// TIA Portal V18 export
// export: Created 2026-11-18T07:26:10.6281665Z, ExportSetting WithDefaults, DisplayName Totally Integrated Automation Portal, DisplayVersion V18 Update 6, DisplayName TIA Portal Openness, DisplayVersion V18 Update 6, DisplayName TIA Portal Version Control Interface, DisplayVersion V18, DisplayName SINAMICS Startdrive Advanced, DisplayVersion V18 SP2 Update 1, DisplayName SINAMICS DCC, DisplayVersion V18 Update 1, DisplayName SINAMICS Startdrive G110M, G120, G120C, G120D, G120P, G115D, DisplayVersion V18 SP2 Update 1, DisplayName SINAMICS Startdrive G130, G150, S120, S150, SINAMICS MV, S210, G220, S200, DisplayVersion V18 SP2 Update 1, DisplayName STEP 7 Professional, DisplayVersion V18 Update 6, DisplayName STEP 7 CFC, DisplayVersion V18 Update 2, DisplayName STEP 7 Safety, DisplayVersion V18, DisplayName WinCC Professional, DisplayVersion V18 Update 6
PlcWatchTable "Drive_1_Izleme"
  PlcWatchTableEntry ""Motor1_Start""  DisplayFormat=Bool, ModifyTrigger=Permanent, MonitorTrigger=Permanent, Comment="Senaryo: start komutu"
  PlcWatchTableEntry ""Motor1_Hiz""  DisplayFormat=DEC_signed, ModifyTrigger=Permanent, MonitorTrigger=Permanent, Comment="Senaryo: hız referansı (rpm)"
  PlcWatchTableEntry ""Motor1_Calisiyor""  DisplayFormat=Bool, ModifyTrigger=Permanent, MonitorTrigger=Permanent, Comment="Senaryo: çalışıyor geri bildirimi"
  PlcWatchTableEntry ""DB_Drive_1_Durum".Calisiyor"  DisplayFormat=Bool, ModifyTrigger=Permanent, MonitorTrigger=Permanent, Comment="Drive_1 çalışıyor (SINA_SPEED AxisEnabled)"
  PlcWatchTableEntry ""DB_Drive_1_Durum".Hata"  DisplayFormat=Bool, ModifyTrigger=Permanent, MonitorTrigger=Permanent, Comment="Drive_1 hata"
  PlcWatchTableEntry ""DB_Drive_1_Durum".Kilit"  DisplayFormat=Bool, ModifyTrigger=Permanent, MonitorTrigger=Permanent, Comment="Drive_1 devreye alma kilidi"
  PlcWatchTableEntry ""DB_Drive_1_Durum".Status"  DisplayFormat=Hex, ModifyTrigger=Permanent, MonitorTrigger=Permanent, Comment="SINA_SPEED Status kelimesi"
  PlcWatchTableEntry ""DB_Drive_1_Durum".Hiz_rpm"  DisplayFormat=Float, ModifyTrigger=Permanent, MonitorTrigger=Permanent, Comment="Gerçek hız (rpm)"
  PlcWatchTableEntry ""DB_Drive_1_Durum".Akim_A"  DisplayFormat=Float, ModifyTrigger=Permanent, MonitorTrigger=Permanent, Comment="Motor akımı (A) = ham / 16384 * Ref_Akim_A"
  PlcWatchTableEntry ""Drive_1_Akim_Ham""  DisplayFormat=DEC_signed, ModifyTrigger=Permanent, MonitorTrigger=Permanent, Comment="Telegram 20 ham akım (IAIST_GLATT, 16384 = %100)"
  PlcWatchTableEntry ""DB_Drive_1_Durum".Tork_Nm"  DisplayFormat=Float, ModifyTrigger=Permanent, MonitorTrigger=Permanent, Comment="Tork (Nm)"
  PlcWatchTableEntry ""DB_Drive_1_Durum".Guc_kW"  DisplayFormat=Float, ModifyTrigger=Permanent, MonitorTrigger=Permanent, Comment="Güç (kW)"
